Fanuc KAREL source: kt00859.KL

-- PROVISIONAL review KL for V770-1; original PC SHA256 6987c1a5ef513ab903bea8d92d49c5bb56ab03f30657415ffa50823e77d22d5c
-- Incomplete behavior may be omitted. Consult companion uncertainty JSON. Do not deploy.
PROGRAM KT00859
%NOLOCKGROUP
VAR
  R1 : REAL
  R2 : REAL
  OUT : REAL
BEGIN
  -- UNRESOLVED_PC offsets 5-16; opcodes 2E,23
  -- UNRESOLVED_PC offsets 21-32; opcodes 2E,23
  -- UNRESOLVED_PC offsets 37-48; opcodes 2E,23
  -- UNRESOLVED_PC offsets 53-64; opcodes 2E,23
  -- UNRESOLVED_PC offsets 69-85; opcodes 27,22,76,64,23
  -- UNRESOLVED_PC offsets 90-94; opcodes 7F
END KT00859
